(* IEC 61131-3 sources: llm-plc-st-eval/data/processed_definitivo/gemini-3.1-pro-preview/B4/zero_shot, 3 files *)

(* ---- ejec_1.st ---- *)
FUNCTION_BLOCK FB_Giro
VAR_INPUT
    btnFwd  : BOOL; // Botón para iniciar giro en sentido horario
    btnRev  : BOOL; // Botón para iniciar giro en sentido antihorario
    btnParo : BOOL; // Botón de paro (TRUE = detener motor)
END_VAR

VAR_OUTPUT
    fwd : BOOL; // Comando de salida para giro horario
    rev : BOOL; // Comando de salida para giro antihorario
END_VAR

(*
   Lógica de control de giro:
   - Se utiliza un circuito de auto-retención (enclavamiento) para cada sentido.
   - La condición "NOT rev" en fwd y "NOT fwd" en rev garantiza que nunca
     estén activas simultáneamente.
   - Al estar enclavado un sentido, presionar el botón del sentido opuesto
     no tendrá efecto. Es obligatorio presionar btnParo primero.
*)

fwd := (btnFwd OR fwd) AND NOT rev AND NOT btnParo;
rev := (btnRev OR rev) AND NOT fwd AND NOT btnParo;

END_FUNCTION_BLOCK

(* ---- ejec_2.st ---- *)
FUNCTION_BLOCK FB_Giro
VAR_INPUT
    btnFwd  : BOOL; // Botón para giro en sentido horario
    btnRev  : BOOL; // Botón para giro en sentido antihorario
    btnParo : BOOL; // Botón de paro (prioridad a la desconexión)
END_VAR

VAR_OUTPUT
    fwd : BOOL; // Salida para motor en sentido horario
    rev : BOOL; // Salida para motor en sentido antihorario
END_VAR

(*
   Lógica de control:
   - NOT btnParo: El paro tiene prioridad absoluta.
   - NOT rev / NOT fwd: Enclavamiento para evitar activación simultánea y obligar a pasar por paro.
   - NOT btnRev / NOT btnFwd: Evita problemas si se pulsan ambos botones a la vez estando el motor detenido.
   - (btnFwd OR fwd): Auto-retención (enclavamiento) de la señal.
*)

fwd := NOT btnParo AND NOT rev AND NOT btnRev AND (btnFwd OR fwd);
rev := NOT btnParo AND NOT fwd AND NOT btnFwd AND (btnRev OR rev);

END_FUNCTION_BLOCK

(* ---- ejec_3.st ---- *)
FUNCTION_BLOCK FB_Giro
VAR_INPUT
    btnFwd  : BOOL; // Botón para iniciar giro en sentido horario
    btnRev  : BOOL; // Botón para iniciar giro en sentido antihorario
    btnParo : BOOL; // Botón de paro (TRUE = detener motor)
END_VAR

VAR_OUTPUT
    fwd : BOOL; // Salida para giro en sentido horario
    rev : BOOL; // Salida para giro en sentido antihorario
END_VAR

(*
   Lógica de giro horario (fwd):
   Se activa con btnFwd o se mantiene enclavada con su propio estado (fwd).
   Condiciones de bloqueo: NO debe estar activo el giro inverso (NOT rev)
   y NO debe estar presionado el botón de paro (NOT btnParo).
*)
fwd := (btnFwd OR fwd) AND NOT rev AND NOT btnParo;

(*
   Lógica de giro antihorario (rev):
   Se activa con btnRev o se mantiene enclavada con su propio estado (rev).
   Condiciones de bloqueo: NO debe estar activo el giro horario (NOT fwd)
   y NO debe estar presionado el botón de paro (NOT btnParo).
*)
rev := (btnRev OR rev) AND NOT fwd AND NOT btnParo;

END_FUNCTION_BLOCK
